Fanuc KAREL source: KT00919.KL

PROGRAM KT00919
%NOLOCKGROUP
VAR
  I1: INTEGER
  I2: INTEGER
  OUT: INTEGER
BEGIN
  I1 = 2
  I2 = 3
  I1 = 2
  I2 = 3
  OUT = INDEX(I1, I1)
END KT00919
